Fanuc KAREL source: kt00601.KL

-- PROVISIONAL review KL for V770-1; original PC SHA256 d94eb6b8a4675474734da3578e0fb109ea9d9541044641e31b0ae816aea6645f
-- Incomplete behavior may be omitted. Consult companion uncertainty JSON. Do not deploy.
PROGRAM KT00601
%NOLOCKGROUP
VAR
  I1 : INTEGER
  I2 : INTEGER
  OUT : INTEGER
BEGIN
  -- UNRESOLVED_PC offsets 5-16; opcodes 2E,23
  -- UNRESOLVED_PC offsets 21-32; opcodes 2E,23
  -- UNRESOLVED_PC offsets 37-48; opcodes 2E,23
  -- UNRESOLVED_PC offsets 53-64; opcodes 2E,23
  -- UNRESOLVED_PC offsets 69-81; opcodes 21,23
  -- UNRESOLVED_PC offsets 86-90; opcodes 7F
END KT00601
